(*
SPDX-FileCopyrightText: © 2026 Oleksandr Tiutyk <trofimich@gmail.com>
SPDX-License-Identifier: MIT
License: https://opensource.org/license/mit
*)

(*!
<summary>Checks the documented completion observation when OnAfterStop resets the timer.</summary>
<description>
The case executes in one PLC callback with a persistent restart probe and no external resources.
AfterTest prepares the fixture for reuse by the runner.
</description>
*)

{attribute 'no_assign'}
{attribute 'no_explicit_call' := 'do not call this function block directly'}
FUNCTION_BLOCK TimerCompletionCallbackTest EXTENDS TOF_Testing.SingleCycleTest
VAR_STAT
	{attribute 'hide'}
	_ClassName : STRING := __POUNAME();
END_VAR
VAR
	_Timer : TimerRestartProbe(name := "Callback reset");
END_VAR

(*!
<summary>Checks the documented completion observation when OnAfterStop resets the timer.</summary>
*)
METHOD PROTECTED ExecuteTest
_Timer.ResetOnAfterStop := TRUE;
_Timer.Interval := TOF_Core.Times.MIN_VALUE;

IF NOT _Timer.Start() THEN
	RecordFailure(message := "Callback probe must accept Start");
	RETURN;
END_IF

Assert.ThatBool(
	actual := _Timer.State.Running,
	message := "Probe must be RUNNING before the completion callback"
).IsTrue();
_Timer.Execute();
Assert.ThatBool(actual := _Timer.State.Ready, message := "Supported callback Reset must restore READY").IsTrue();
Assert.ThatBool(
	actual := _Timer.Triggered,
	message := "Callback Reset may clear the pulse before Execute returns"
).IsFalse();
Assert.ThatBool(actual := _Timer.Elapsed, message := "Callback Reset must clear retained Q").IsFalse();
Assert.ThatBool(
	actual := _Timer.ElapsedTime = TOF_Core.Times.MIN_VALUE,
	message := "Callback Reset must clear ET"
).IsTrue();
END_METHOD

(*!
<summary>Returns the owned timer to READY before reporting the result.</summary>
<description>
Reopens the stopping gate and disables callback injections before cooperative cleanup.
</description>
*)
METHOD PROTECTED AfterTest
_Timer.AllowStopping := TRUE;
_Timer.ThrowOnBeforeStart := FALSE;
_Timer.ThrowOnReset := FALSE;
_Timer.ResetOnAfterStop := FALSE;

Assert.ThatBool(
	actual := PrepareTimerTestForReuse(timer := _Timer),
	message := "The timer must return to READY after cleanup"
).IsTrue();
END_METHOD

//! <summary>Borrows the concrete class name. Callers must not modify it.</summary>
{attribute 'monitoring' := 'call'}
PROPERTY ClassName : REFERENCE TO STRING
GET
ClassName REF= _ClassName;
END_GET
END_PROPERTY

//! <summary>Borrows the compiler-initialized namespace. Callers must not modify it.</summary>
{attribute 'monitoring' := 'call'}
PROPERTY NamespaceName : REFERENCE TO STRING
GET
NamespaceName REF= CurrentNamespace.Name;
END_GET
END_PROPERTY

//! <summary>Reports the concrete instance size in bytes.</summary>
{attribute 'monitoring' := 'call'}
PROPERTY SelfSize : ULINT
GET
SelfSize := XSIZEOF(THIS^);
END_GET
END_PROPERTY

END_FUNCTION_BLOCK

(* stored: Version 1.1.0.1
   POU TimerCompletionCallbackTest: Id {9c80ffbb-735b-4a83-96b7-985e778a39e4}, SpecialFunc None
   Method ExecuteTest: Id {6aeec917-ee8e-4389-9643-6409fa239964}
   Method AfterTest: Id {6b427096-29c4-4f16-bce6-84f0a6e642c7}
   Property ClassName: Id {982ecb15-2358-495a-8ba2-3d4524b8d938}
   Get Get: Id {54df6790-bdd6-4349-ab5f-887f345ce92b}
   Property NamespaceName: Id {37040404-5e77-4cf3-89ad-75717c971896}
   Get Get: Id {db372d89-dae0-4cce-a1c0-3a17abca6a57}
   Property SelfSize: Id {046c86af-bd45-41b0-9906-6807885678f9}
   Get Get: Id {c41434d4-6ee2-409c-b3ca-b95b79ca204e} *)
